{attribute 'qualified_only'}
VAR_GLOBAL
	bWartungseinheitEntluften		: BOOL;   //MaintenanceUnitVenting
	bLaserEnable					: BOOL;

	bCWTrigger						: BOOL;
	bCWSTO							: BOOL;
	bCWJob							: BOOL;

	bVentilAuswerferAS				: BOOL;   //ValveEjector
	bVentilAuswerferGS				: BOOL;   //ValveEjector
	bVentilSpannerAS				: BOOL;   //ValveClamp
	bVentilSpannerGS				: BOOL;   //ValveClamp
	bVentilWeicheAS					: BOOL;   //ValveDiverter
	bVentilWeicheGS					: BOOL;   //ValveDiverter
	bVentilAusblastenAS				: BOOL;   //BlowOutValve
	bVentilAusblastenGS				: BOOL;   //BlowOutValve	
	
	bVentilEinlaufAS				: BOOL;   //ValveInfeed
	bVentilEinlaufGS				: BOOL;   //ValveInfeed
	bVentilAuslaufAS				: BOOL;   //ValveOutfeed
	bVentilAuslaufGS				: BOOL;   //ValveOutfeed	
	bVentilAuswerfBypassAS			: BOOL;   //EjectionBypassValve
	bVentilAuswerfBypassGS			: BOOL;   //EjectionBypassValve

END_VAR

(* stored: Version 1.1.0.1
   GVL GVL_Outputs: Id {dc412ae4-fcc4-4abc-90fc-9e0d95b76746} *)
